(* IEC 61131-3 sources: Test-Git_ESME26/00_Initial Project_LB.fbsproj/M660.device.xml.v3^/Plc Logic.plclogic.xml.v3^/Application.application.xml.v3^/Global Variables, 1 file *)

(* ---- GVL.gvl ---- *)
{attribute 'qualified_only'}
VAR_GLOBAL
END_VAR
